FUNCTION_BLOCK DEMUX_X3 (* Basic Function Block Type *)
  (* Standard: 61499-2 *)
  (* Version 0.0, 10/11/2026, macie, nxtControl GmBH, Template *)
  PACKAGE Main;
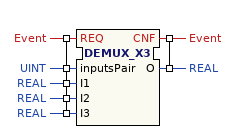
  EVENT_INPUT
    REQ WITH inputsPair, I1, I2, I3; (* Normal Execution Request *)
  END_EVENT
  EVENT_OUTPUT
    CNF WITH O; (* Execution Confirmation *)
  END_EVENT
  VAR_INPUT
    inputsPair : UINT;
    I1 : REAL; (* Input event qualifier *)
    I2 : REAL;
    I3 : REAL;
  END_VAR
  VAR_OUTPUT
    O : REAL; (* Output event qualifier *)
  END_VAR
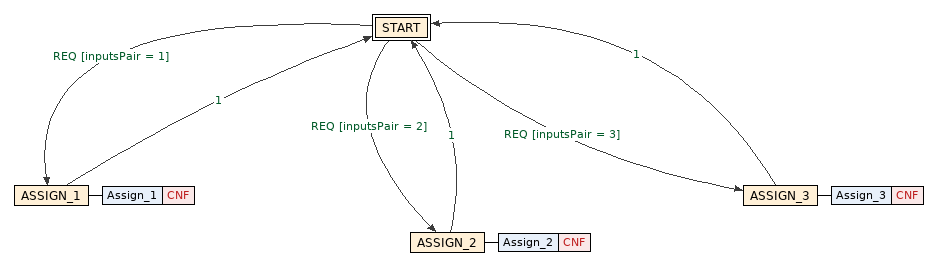
  EC_STATES
    START; (* Initial State *)
    ASSIGN_1 : Assign_1 -> CNF;
    ASSIGN_2 : Assign_2 -> CNF;
    ASSIGN_3 : Assign_3 -> CNF;
  END_STATES
  EC_TRANSITIONS
    START TO ASSIGN_1 := REQ [inputsPair = 1];
    ASSIGN_1 TO START := 1;
    START TO ASSIGN_2 := REQ [inputsPair = 2];
    START TO ASSIGN_3 := REQ [inputsPair = 3];
    ASSIGN_2 TO START := 1;
    ASSIGN_3 TO START := 1;
  END_TRANSITIONS
  ALGORITHM INIT IN ST: (* Initialization algorithm *)
;
  END_ALGORITHM
  ALGORITHM REQ IN ST: (* Normally executed algorithm *)
;
  END_ALGORITHM
  ALGORITHM Assign_1 IN ST:
;
O := I1;
  END_ALGORITHM
  ALGORITHM Assign_2 IN ST:
;
O := I2;
  END_ALGORITHM
  ALGORITHM Assign_3 IN ST:
;
O := I3;
  END_ALGORITHM
END_FUNCTION_BLOCK
